(* CoDeSys 2.3 export: 02_timers_tellers.exp *)
(* Libraries: Standard.lib 2.12.10 14:48:34 *)

(* Global variable list: Globale_Variablen *)
VAR_GLOBAL
	iStart			AT %IX0.0 : BOOL;
	iStop			AT %IX0.1 : BOOL;
	iAtPusher		AT %IX0.2 : BOOL;
	iSimRunning		AT %IX0.6 : BOOL;

	oConveyor		AT %QX0.0 : BOOL;
	oPusher			AT %QX0.1 : BOOL;
	oEmitter		AT %QX0.2 : BOOL;
	oRunLamp		AT %QX0.3 : BOOL;
	wAantal			AT %QW2 : WORD;

	tVerstreken		: TIME;				(* zonder adres: alleen op naam te koppelen *)
END_VAR

(* POU PLC_PRG, ST *)
PROGRAM PLC_PRG
VAR
	bRun			: BOOL;
	tonStart		: TON;		(* vertraagde start van de band *)
	tofNaloop		: TOF;		(* naloop van de lamp *)
	tpPuls			: TP;		(* vaste puls bij elke doos *)
	rtDoos			: R_TRIG;	(* doos komt aan *)
	ftDoos			: F_TRIG;	(* doos vertrekt *)
	ctuDozen		: CTU;		(* dozenteller *)
	ctdRest			: CTD;		(* aftellen tot batch klaar *)
	srFout			: SR;
	bBatchKlaar		: BOOL;
END_VAR
IF iStop OR NOT iSimRunning THEN
	bRun := FALSE;
ELSIF iStart THEN
	bRun := TRUE;
END_IF;

(* Band start 2 s na het startcommando *)
tonStart(IN := bRun, PT := T#2s);

(* Flanken van de photo-eye *)
rtDoos(CLK := iAtPusher);
ftDoos(CLK := iAtPusher);

(* Tellen: omhoog per aangekomen doos, reset met stop *)
ctuDozen(CU := rtDoos.Q, RESET := iStop, PV := 10);
ctdRest(CD := ftDoos.Q, LOAD := iStart, PV := 5);
bBatchKlaar := ctdRest.Q;

(* Puls van 500 ms bij elke doos, lamp met 1 s naloop *)
tpPuls(IN := rtDoos.Q, PT := T#500ms);
tofNaloop(IN := bRun, PT := T#1s);

(* Fout: tien dozen geteld zonder stop *)
srFout(SET1 := ctuDozen.Q, RESET := iStop);

oConveyor := tonStart.Q AND NOT srFout.Q1;
oEmitter := tonStart.Q AND NOT bBatchKlaar;
oPusher := tpPuls.Q;
oRunLamp := tofNaloop.Q;
wAantal := INT_TO_WORD(ctuDozen.CV);
tVerstreken := tonStart.ET;
END_PROGRAM
